// TIA Portal V21 export
// export: Created 2026-08-21T20:18:56.8671985Z, ExportSetting None, DisplayName Totally Integrated Automation Portal, DisplayVersion V21, DisplayName STEP 7 Professional, DisplayVersion V21, DisplayName STEP 7 Safety, DisplayVersion V21, DisplayName Tech WebApplication, DisplayVersion V21, DisplayName WinCC Basic/Comfort/Advanced, DisplayVersion V21, DisplayName WinCC Professional, DisplayVersion V21, DisplayName WinCC Unified, DisplayVersion V21
TYPE "UDT_Service_ProcedureRawDataMedium"
   STRUCT
      procedure { S7_SetPoint := 'True'} : Array[0..15] of "UDT_MTP_ProcedureExtended";
   END_STRUCT;
END_TYPE
